TYPE ST_Config :
STRUCT
    speed : T_Speed;
    delay : TIME := T#100ms;
    enabled : BOOL := TRUE;
END_STRUCT
END_TYPE

(* stored: Version 1.1.0.1 *)
